(* IEC 61131-3 sources: iolistgen/tools/tests/fixtures/sourcemap/src/DUTs, 2 files *)

(* ---- ST_Probe.dut.st ---- *)
// Многострочные начальное значение массива и вложенный массив в полях структуры
TYPE ST_Probe :
STRUCT
    arStep : ARRAY[1..4] OF REAL := [0.5, 1.0,
        1.5, 2.0];
    aaiGrid : ARRAY[0..1] OF
        ARRAY[0..2] OF INT;
    sName : STRING(GVL_Const.NAME_SIZE) := 'abc';   // @8
    rLim : REAL := 1.0;                               // @9
END_STRUCT
END_TYPE

(* ---- T_Percent.dut.st ---- *)
// Псевдоним с поддиапазоном: начальное значение вне диапазона — OutOfBounds iec_checker
TYPE T_Percent : INT(0..100) := 200;
END_TYPE
